// CFC twin of T_SafeEdm_Tests: the same tests drawn as CFC diagrams, the way a TwinSAFE project is authored.
    FUNCTION_BLOCK T_SafeEdm_Tests_CFC EXTENDS T_SafeCfcTestSuite
    VAR
    // Test_SwitchOnTimeoutGivesError
    group_1 : T_SafeGroup;
    fb_1 : T_SafeEdm(group := group_1) := (Parameters := (SwitchOnTime := T#100MS));
    t1_1 : TON;
    trig1_1 : R_TRIG;
    // Test_NoErrorWhenFeedbackFollows
    group_2 : T_SafeGroup;
    fb_2 : T_SafeEdm(group := group_2) := (Parameters := (SwitchOnTime := T#100MS, SwitchOffTime := T#100MS));
    t1_2 : TON;
    t2_2 : TON;
    trig1_2 : R_TRIG;
    trig2_2 : R_TRIG;
END_VAR

Test_SwitchOnTimeoutGivesError();
Test_NoErrorWhenFeedbackFollows();

METHOD PRIVATE Test_SwitchOnTimeoutGivesError
// note: this text did not pass the execution check against the stored diagram
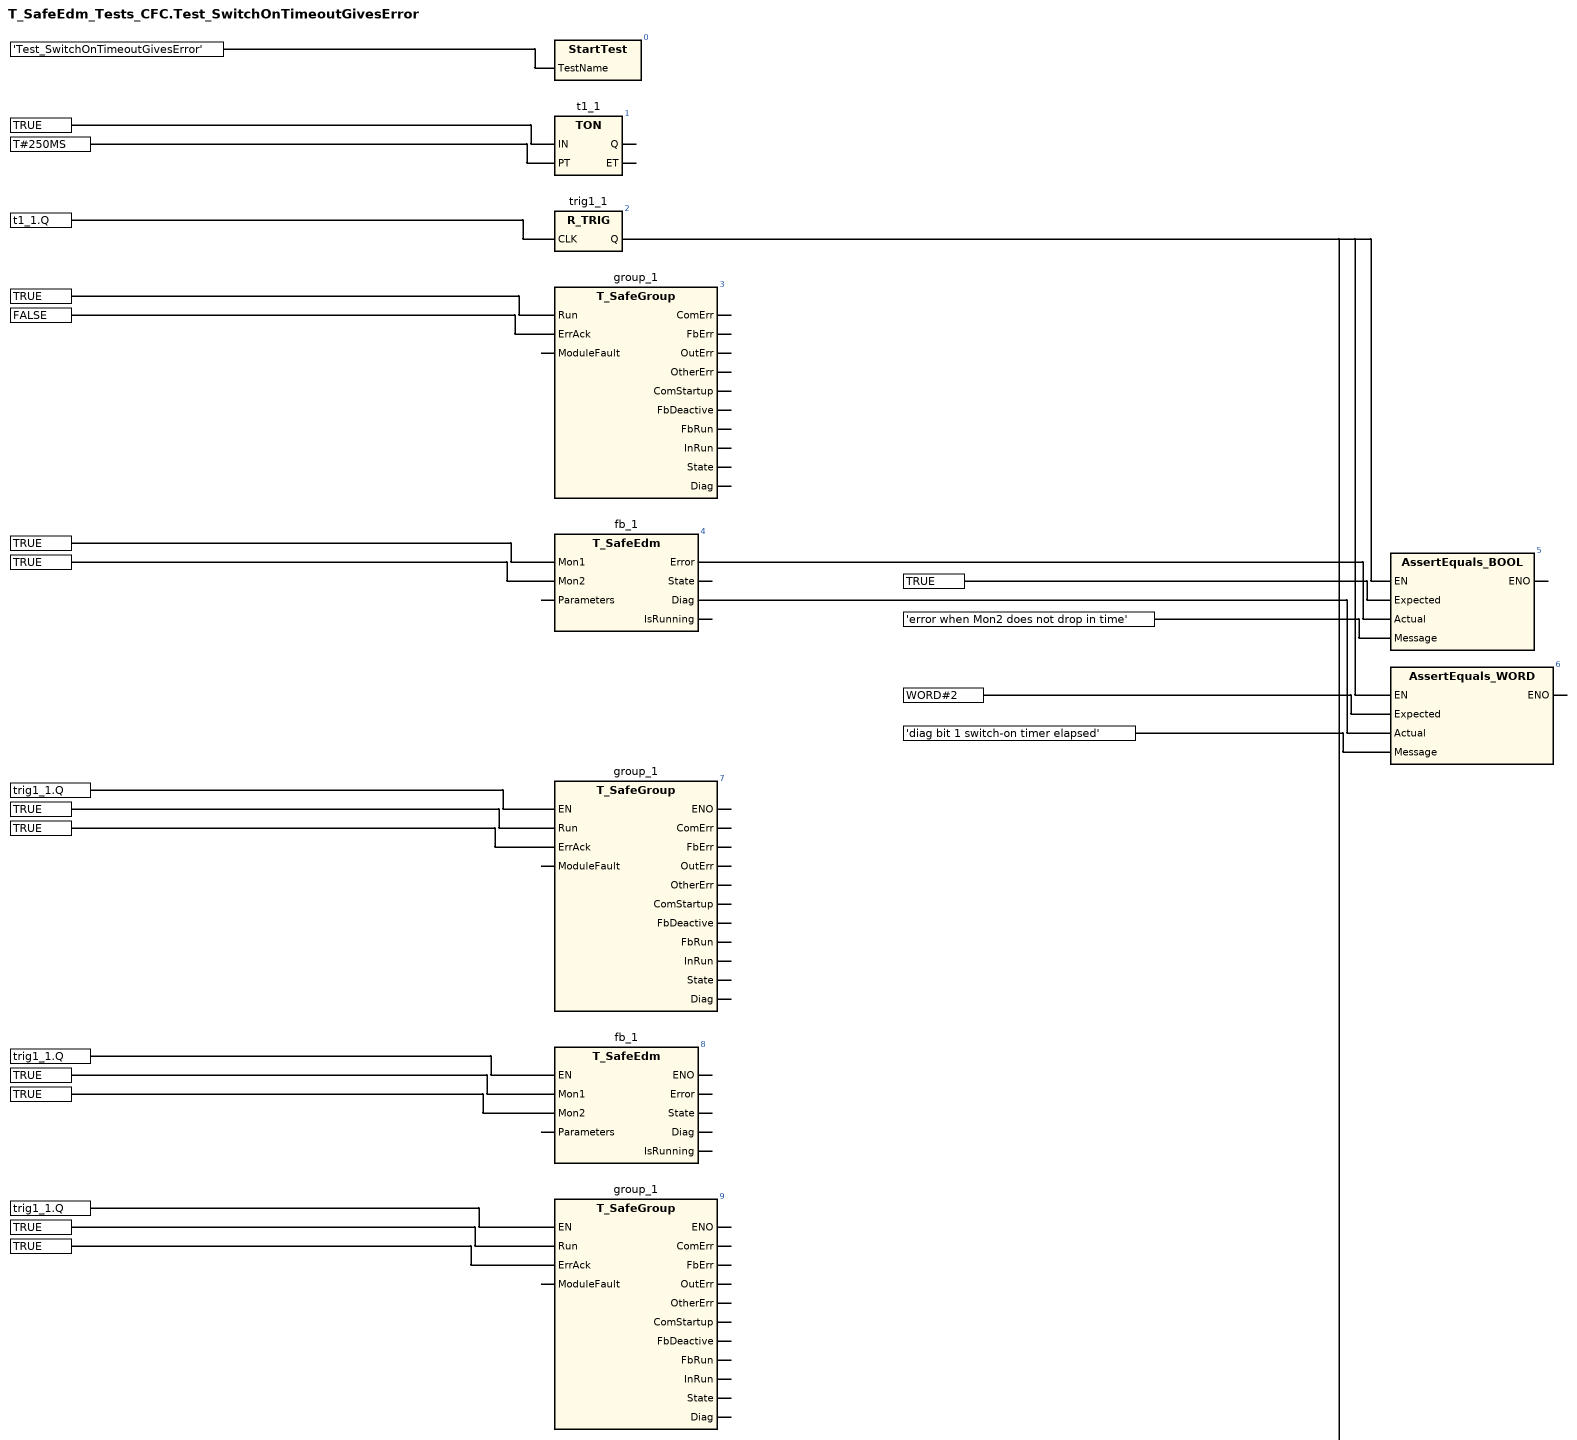
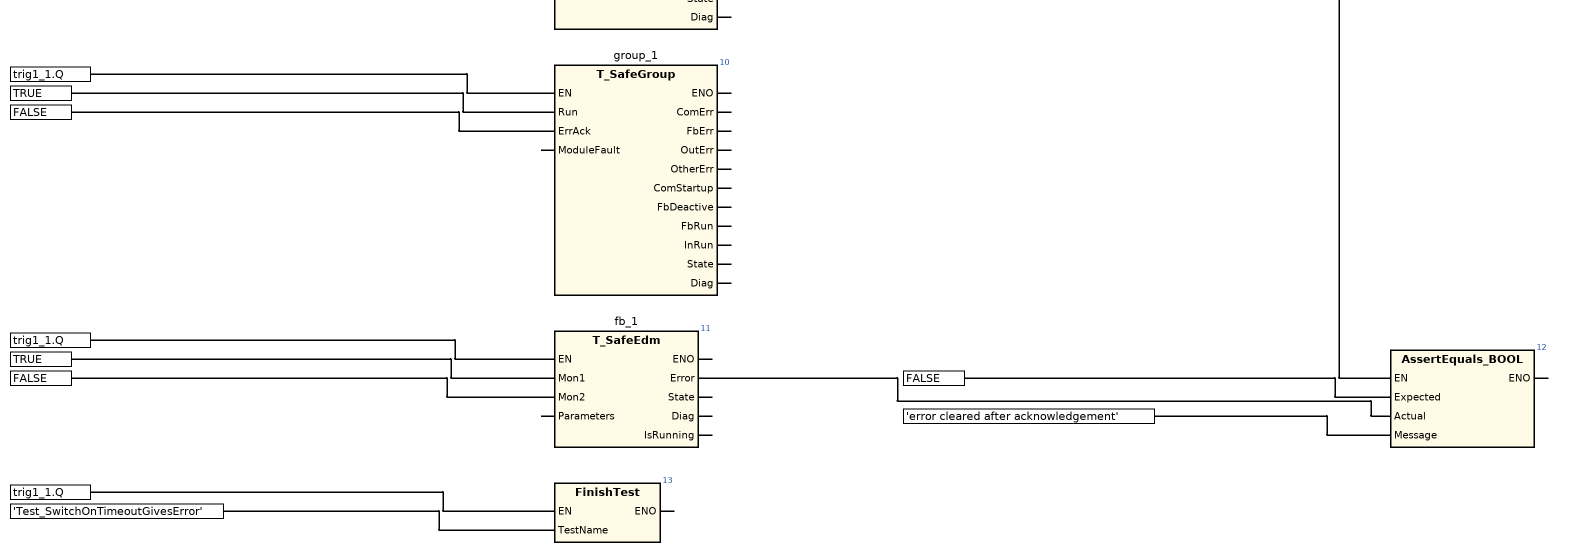
StartTest(TestName := 'Test_SwitchOnTimeoutGivesError');
t1_1(IN := TRUE, PT := T#250MS); // TON
trig1_1(CLK := t1_1.Q); // R_TRIG
group_1(Run := TRUE, ErrAck := FALSE); // T_SafeGroup
fb_1(Mon1 := TRUE, Mon2 := TRUE); // T_SafeEdm
IF trig1_1.Q THEN AssertEquals_BOOL(Expected := TRUE, Actual := fb_1.Error, Message := 'error when Mon2 does not drop in time'); END_IF
IF trig1_1.Q THEN AssertEquals_WORD(Expected := WORD#2, Actual := fb_1.Diag, Message := 'diag bit 1 switch-on timer elapsed'); END_IF
IF trig1_1.Q THEN
    group_1(Run := TRUE, ErrAck := TRUE); // T_SafeGroup
END_IF
IF trig1_1.Q THEN
    fb_1(Mon1 := TRUE, Mon2 := TRUE); // T_SafeEdm
END_IF
IF trig1_1.Q THEN
    group_1(Run := TRUE, ErrAck := TRUE); // T_SafeGroup
END_IF
IF trig1_1.Q THEN
    group_1(Run := TRUE, ErrAck := FALSE); // T_SafeGroup
END_IF
IF trig1_1.Q THEN
    fb_1(Mon1 := TRUE, Mon2 := FALSE); // T_SafeEdm
END_IF
IF trig1_1.Q THEN AssertEquals_BOOL(Expected := FALSE, Actual := fb_1.Error, Message := 'error cleared after acknowledgement'); END_IF
IF trig1_1.Q THEN FinishTest(TestName := 'Test_SwitchOnTimeoutGivesError'); END_IF
END_METHOD

METHOD PRIVATE Test_NoErrorWhenFeedbackFollows
// note: this text did not pass the execution check against the stored diagram
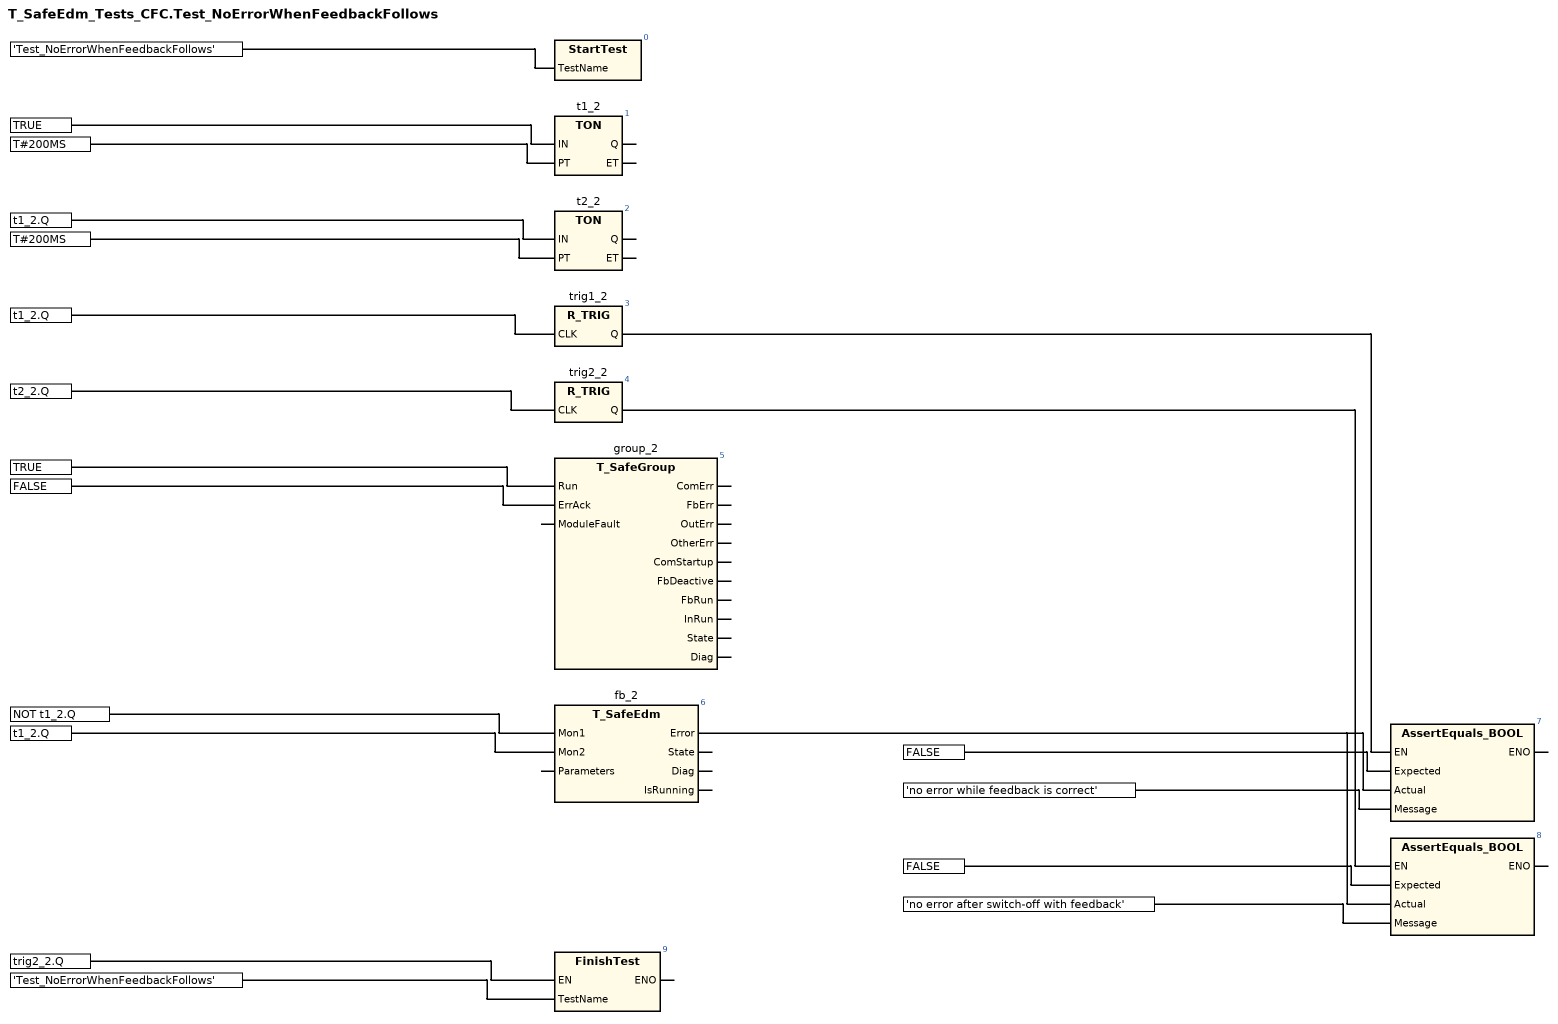
StartTest(TestName := 'Test_NoErrorWhenFeedbackFollows');
t1_2(IN := TRUE, PT := T#200MS); // TON
t2_2(IN := t1_2.Q, PT := T#200MS); // TON
trig1_2(CLK := t1_2.Q); // R_TRIG
trig2_2(CLK := t2_2.Q); // R_TRIG
group_2(Run := TRUE, ErrAck := FALSE); // T_SafeGroup
fb_2(Mon1 := NOT t1_2.Q, Mon2 := t1_2.Q); // T_SafeEdm
IF trig1_2.Q THEN AssertEquals_BOOL(Expected := FALSE, Actual := fb_2.Error, Message := 'no error while feedback is correct'); END_IF
IF trig2_2.Q THEN AssertEquals_BOOL(Expected := FALSE, Actual := fb_2.Error, Message := 'no error after switch-off with feedback'); END_IF
IF trig2_2.Q THEN FinishTest(TestName := 'Test_NoErrorWhenFeedbackFollows'); END_IF
END_METHOD

END_FUNCTION_BLOCK

(* stored: Version 1.1.0.1, ProductVersion 3.1.4026.22
   POU T_SafeEdm_Tests_CFC: Id {8b16f178-cc2a-5f1f-a536-cb9a23f0b9b3}, SpecialFunc None
   Method Test_SwitchOnTimeoutGivesError: Id {c7b4d270-31ce-5f50-8fda-118c2e6518c2}
   Method Test_NoErrorWhenFeedbackFollows: Id {8d4290d6-3027-5731-bab7-d393c6d99d61} *)
